(* IEC 61131-3 sources: Lasal-MCP/examples/SampleSource/4_PumpControlSchemeSolution/Stations/MachineControl/MachineControl/Class/ButtonStates, 1 file *)

(* ---- ButtonStates.st ---- *)
(*!
<Class
	Name               = "ButtonStates"
	Revision           = "0.0"
	RealtimeTask       = "false"
	CyclicTask         = "false"
	BackgroundTask     = "false"
	Sigmatek           = "false"
	OSInterface        = "false"
	HighPriority       = "false"
	Automatic          = "false"
	UpdateMode         = "Prescan"
	SharedCommandTable = "true"
	Objectsize         = "(496,0)">
	<Channels>
		<Server Name="DataSvrScheme" Visualized="true" Initialize="false" WriteProtected="false" Retentive="false"/>
		<Server Name="ObjectScheme" Visualized="true" Initialize="false" WriteProtected="false" Retentive="false"/>
		<Server Name="UnitScheme" Visualized="true" Initialize="false" WriteProtected="false" Retentive="false"/>
	</Channels>
</Class>
*)
ButtonStates : CLASS
  //Servers:
	UnitScheme 	: SvrChCmd_DINT;
	DataSvrScheme 	: SvrCh_DINT;
	ObjectScheme 	: SvrCh_DINT;
  //Clients:
  //Variables:
  //Functions:
  //Tables:
	FUNCTION @STD
		VAR_OUTPUT
			ret_code	: CONFSTATES;
		END_VAR;
	FUNCTION GLOBAL TAB @CT_;
END_CLASS;
